Staubli VAL3: ifItem.pjx

--- ifItem.pjx ---
Parameters version=s8.10.3Cs9_BS2093 stackSize=5000 millimeterUnit=true
Program file=start.pgx
Program file=stop.pgx
Data file=ifItem.dtx

--- ifItem.dtx ---
public num nSigType[3]
public num nSigIndex[3]
public num nValue[3]
public bool bANDOR[2]

--- start.pgx ---
program start()
begin
end

--- stop.pgx ---
program stop()
begin
end
